// TIA Portal V21 export
VAR_GLOBAL   // PLC tag table "EIO_Odot"
   A1 AT %I8.0 : Bool;   // Pnematik Endlagenschalter B1
   A2 AT %I8.1 : Bool;   // Pnematik Endlagenschalter B2
   B1 AT %I8.2 : Bool;
   B2 AT %I8.3 : Bool;
   di_Warenträger AT %I10.0 : Bool;   // Warenträger erkannt
   di_einschubachse_ref AT %I10.1 : Bool;   // Referenzierung für z-Einschub
   di_EnableXYMovement AT %I10.2 : Bool;   // Sensor für erkennen ob z-Einschub eingefahren ist. Horizontale und Vertikale Achse dürfen nur fahren wenn dieser Sensor =0 ist!
   "A" AT %Q4.0 : Bool;   // Pnematikzylinder B
   "B" AT %Q4.1 : Bool;
   Notaus_IO AT %Q4.7 : Bool;
END_VAR
